// assert
AssertEquals_BOOL(Expected := TRUE, Actual := terminal_2.Channel1, Message := 'Channel1 follows SafeOut1');
AssertEquals_BOOL(Expected := FALSE, Actual := terminal_2.Channel2, Message := 'Channel2 follows SafeOut2');

// act: swap
group_2(Run := TRUE);
terminal_2(SafeOut1 := FALSE, SafeOut2 := TRUE, StartupTime := T#0S);

// assert
AssertEquals_BOOL(Expected := FALSE, Actual := terminal_2.Channel1, Message := 'Channel1 swapped');
AssertEquals_BOOL(Expected := TRUE, Actual := terminal_2.Channel2, Message := 'Channel2 swapped');
TEST_FINISHED_NAMED(__POUNAME());
END_METHOD

METHOD PRIVATE Test_ComErrorForcesChannelsFalse
TcUnit.TEST(__POUNAME());

// arrange: in Data with both outputs on
FOR i_3 := 1 TO 5 DO
    group_3(Run := TRUE);
    terminal_3(SafeOut1 := TRUE, SafeOut2 := TRUE, StartupTime := T#0S);
END_FOR
AssertEquals_BOOL(Expected := TRUE, Actual := terminal_3.Channel2, Message := 'Channel2 on before the error');

// act
group_3(Run := TRUE);
terminal_3(SafeOut1 := TRUE, SafeOut2 := TRUE, InjectComError := TRUE, StartupTime := T#0S);

// assert
AssertEquals_BOOL(Expected := TRUE, Actual := terminal_3.ComError, Message := 'com error');
AssertEquals_BOOL(Expected := FALSE, Actual := terminal_3.Channel1, Message := 'Channel1 fail-safe on com error');
AssertEquals_BOOL(Expected := FALSE, Actual := terminal_3.Channel2, Message := 'Channel2 fail-safe on com error');
TEST_FINISHED_NAMED(__POUNAME());
END_METHOD

METHOD PRIVATE Test_RegistersAsConnection
TcUnit.TEST(__POUNAME());

// act
group_4(Run := TRUE);
terminal_4(StartupTime := T#0S);

// assert
AssertEquals_UINT(Expected := 1, Actual := group_4.ConnectionCount, Message := 'one connection registered');
AssertEquals_UINT(Expected := 0, Actual := group_4.FunctionBlockCount, Message := 'no function blocks');
TEST_FINISHED_NAMED(__POUNAME());
END_METHOD

METHOD PRIVATE Test_GroupNotRunningForcesChannelsFalse
TcUnit.TEST(__POUNAME());
// arrange: connection in Data with the group running
FOR i_5 := 1 TO 10 DO
    group_5(Run := TRUE, ModuleFault := FALSE);
    terminal_5(StartupTime := T#0S, SafeOut1 := TRUE, SafeOut2 := TRUE);
END_FOR
AssertEquals_BOOL(Expected := TRUE, Actual := terminal_5.Channel1, Message := 'channel on while the group runs');
// act: group STOP (the connection stays in Data)
group_5(Run := FALSE, ModuleFault := FALSE);
terminal_5(StartupTime := T#0S, SafeOut1 := TRUE, SafeOut2 := TRUE);
// assert
AssertEquals_BOOL(Expected := TRUE, Actual := terminal_5.InDataState, Message := 'still in Data');
AssertEquals_BOOL(Expected := FALSE, Actual := terminal_5.Channel1, Message := 'outputs off with the group in STOP');
// act: group ERROR
group_5(Run := TRUE, ModuleFault := TRUE);
terminal_5(StartupTime := T#0S, SafeOut1 := TRUE, SafeOut2 := TRUE);
group_5(Run := TRUE, ModuleFault := TRUE);
terminal_5(StartupTime := T#0S, SafeOut1 := TRUE, SafeOut2 := TRUE);
AssertEquals_BYTE(Expected := TO_BYTE(E_SafeGroupState.Error), Actual := group_5.State, Message := 'group in ERROR');
AssertEquals_BOOL(Expected := FALSE, Actual := terminal_5.Channel2, Message := 'outputs off with the group in ERROR');
TEST_FINISHED_NAMED(__POUNAME());
END_METHOD

END_FUNCTION_BLOCK

// ---- Core/T_SafeOutputTerminal2.TcPOU
// Model of a two channel safe output terminal (EL2912): a TwinSAFE connection with two channels.
// Declare it in its group:  outputTerminal : T_SafeOutputTerminal2(group := safetyGroup);
// SafeOut1..2 are wired from FB outputs; Channel1..2 are the simulated field outputs,
// forced FALSE (fail-safe) unless the connection is in the Data state and the group is in RUN (OutputsEnabled).
FUNCTION_BLOCK T_SafeOutputTerminal2 EXTENDS T_SafeConnection
VAR_INPUT
    SafeOut1 : BOOL;
    SafeOut2 : BOOL;
END_VAR
VAR_OUTPUT
    Channel1 : BOOL;
    Channel2 : BOOL;
END_VAR

SUPER^();
Channel1 := SafeOut1 AND OutputsEnabled;
Channel2 := SafeOut2 AND OutputsEnabled;

END_FUNCTION_BLOCK

// ---- Tests/T_SafeConnShutdown_Tests.TcPOU
FUNCTION_BLOCK T_SafeConnShutdown_Tests EXTENDS TcUnit.FB_TestSuite
VAR
    // Test_DeactivateShutsDownConnection
    group_1 : T_SafeGroup;
    conn_1 : T_SafeConnection(group := group_1);
    fb_1 : T_SafeConnShutdown(group := group_1, connection := conn_1);
    i_1 : INT;
END_VAR

Test_DeactivateShutsDownConnection();

METHOD PRIVATE Test_DeactivateShutsDownConnection
TcUnit.TEST(__POUNAME());

// arrange: connection up
FOR i_1 := 1 TO 5 DO
    group_1(Run := TRUE);
    conn_1(StartupTime := T#0S);
    fb_1(Deactivate1 := FALSE);
END_FOR

AssertEquals_BOOL(Expected := FALSE, Actual := fb_1.Deactivated, Message := 'connection up');
// act
group_1(Run := TRUE);
fb_1(Deactivate1 := TRUE);
conn_1(StartupTime := T#0S);
fb_1(Deactivate1 := TRUE);
// assert
AssertEquals_BOOL(Expected := TRUE, Actual := conn_1.IsShutdown, Message := 'connection shut down');
AssertEquals_BOOL(Expected := TRUE, Actual := fb_1.Deactivated, Message := 'Deactivated output on');

// act: release
FOR i_1 := 1 TO 6 DO
    group_1(Run := TRUE);
    fb_1(Deactivate1 := FALSE);
    conn_1(StartupTime := T#0S);
END_FOR

AssertEquals_BOOL(Expected := TRUE, Actual := conn_1.InDataState, Message := 'connection re-established');
AssertEquals_BOOL(Expected := FALSE, Actual := fb_1.Deactivated, Message := 'Deactivated output off');
TEST_FINISHED_NAMED(__POUNAME());
END_METHOD

END_FUNCTION_BLOCK

// ---- FunctionBlocks/T_SafeConnShutdown.TcPOU
// Model of the TwinSAFE FB CONNECTION SHUTDOWN.
// Shuts down the assigned connection while the Deactivate inputs are TRUE and reports Deactivated
// once the connection is shut down (also when the partner shut it down). The connection is assigned
// at construction (the Connection ID of the Safety Editor):
//     connShutdown : T_SafeConnShutdown(group := safetyGroup, connection := toolConnection);
{attribute 'reflection'}
FUNCTION_BLOCK T_SafeConnShutdown EXTENDS T_SafeFunctionBlockBase
VAR_INPUT
    Deactivate1 : BOOL;
    Deactivate2 : BOOL;
    Parameters : ST_SafeConnShutdownParameters;
END_VAR
VAR_OUTPUT
    Deactivated : BOOL;
END_VAR
VAR
    {attribute 'is_connected' := 'Deactivate1'}
    _deactivate1Connected : BOOL;
    {attribute 'is_connected' := 'Deactivate2'}
    _deactivate2Connected : BOOL;
    _connection : REFERENCE TO T_SafeConnection;
    _pairs : ARRAY[1..1] OF T_SafeInputPair;
    _state : E_SafeFbState := E_SafeFbState.Stop;
    _prevState : E_SafeFbState;
END_VAR

SUPER^();

PROPERTY ConnShutdownState : E_SafeFbState
GET
ConnShutdownState := _state;
END_GET
END_PROPERTY

METHOD FB_init : BOOL
VAR_INPUT
    bInitRetains : BOOL;
    bInCopyCode : BOOL;
    group : REFERENCE TO T_SafeGroup; // the TwinSAFE group this block belongs to
    connection : REFERENCE TO T_SafeConnection; // the connection to shut down (Connection ID)
END_VAR
// the base FB_init (group registration) is called implicitly by TwinCAT
_connection REF= connection;
END_METHOD

METHOD PROTECTED Process
VAR
    acknowledge : BOOL;
    deactivate : BOOL;
    operating : BOOL;
    stateBefore : E_SafeFbState;
    passes : USINT;
END_VAR
acknowledge := (_state = E_SafeFbState.Error) AND _errAck;
_pairs[1](
    In1 := Deactivate1,
    In2 := Deactivate2,
    Active1 := _deactivate1Connected,
    Active2 := _deactivate2Connected,
    MakeContact1 := Parameters.Deactivate1MakeContact,
    MakeContact2 := Parameters.Deactivate2MakeContact,
    DiscrepancyTime := Parameters.DiscrepancyTime,
    Monitor := _fbRun,
    SafeInputsAfterDiscError := Parameters.SafeInputsAfterDiscError,
    Acknowledge := acknowledge
);

deactivate := _pairs[1].IsActive AND _pairs[1].AllTrue;

IF NOT _fbRun AND _state <> E_SafeFbState.Error AND _state <> E_SafeFbState.Reset THEN
    _state := E_SafeFbState.Stop;
END_IF

operating := (_state = E_SafeFbState.Safe) OR (_state = E_SafeFbState.Run);

IF _pairs[1].DiscrepancyError AND operating THEN
    UpdateDiscrepancyDiag();
    _state := E_SafeFbState.Error;
END_IF

passes := 0;

REPEAT
    stateBefore := _state;

    CASE _state OF
        E_SafeFbState.Stop:
            IF StateChanged() THEN
                Deactivated := FALSE;
                Error       := FALSE;
                Diag        := 0;
            END_IF

            _connection.LocalShutdown := FALSE;

            IF _fbRun THEN
                _state := E_SafeFbState.Safe;
            END_IF

        E_SafeFbState.Safe:
            IF StateChanged() THEN
                Deactivated := FALSE;
            END_IF

            _connection.LocalShutdown := deactivate;

            IF _connection.IsShutdown THEN
                _state := E_SafeFbState.Run;
            END_IF

        E_SafeFbState.Run:
            IF StateChanged() THEN
                Deactivated := TRUE;
            END_IF

            _connection.LocalShutdown := deactivate;

            IF NOT _connection.IsShutdown THEN
                _state := E_SafeFbState.Safe;
            END_IF

        E_SafeFbState.Error:
            IF StateChanged() THEN
                Deactivated := FALSE;
                Error       := TRUE;
            END_IF

            _connection.LocalShutdown := FALSE;
            UpdateDiscrepancyDiag();

            IF _errAck AND NOT _pairs[1].DiscrepancyError THEN
                _state := E_SafeFbState.Reset;
            END_IF

        E_SafeFbState.Reset:
            IF StateChanged() THEN
                Error := FALSE;
                Diag  := 0;
            END_IF

            IF _errAckFallingEdge THEN
                _state := SEL(_fbRun, E_SafeFbState.Stop, E_SafeFbState.Safe);
            END_IF
    END_CASE

    passes := passes + 1;
UNTIL (stateBefore = _state) OR (passes >= 3)
END_REPEAT

State := TO_BYTE(_state);
END_METHOD

METHOD PRIVATE StateChanged : BOOL
IF _prevState = _state THEN
    RETURN;
END_IF

_prevState   := _state;
StateChanged := TRUE;
END_METHOD

// Mirrors the discrepancy state of every pair into the diagnostic bits.
METHOD PRIVATE UpdateDiscrepancyDiag
VAR
    i : USINT;
END_VAR
FOR i := 1 TO 1 DO
    IF _pairs[i].DiscrepancyError THEN
        SetDiagBit(0);

        IF _pairs[i].AwaitingSafeInputs THEN
            SetDiagBit(8);
        ELSE
            ClearDiagBit(8);
        END_IF
    END_IF
END_FOR
END_METHOD

END_FUNCTION_BLOCK

// ---- Tests/T_SafeGroup_Tests.TcPOU
FUNCTION_BLOCK T_SafeGroup_Tests EXTENDS TcUnit.FB_TestSuite
VAR
    // Test_StopWhenRunFalse
    group_1 : T_SafeGroup;
    fb_1 : T_SafeAnd(group := group_1);
    // Test_RunsFunctionBlocksWithoutConnections
    group_2 : T_SafeGroup;
    fb_2 : T_SafeAnd(group := group_2);
    // Test_FbErrorStopsGroupAndErrAckRecovers
    group_3 : T_SafeGroup;
    eStop_3 : T_SafeEStop(group := group_3);
    andFb_3 : T_SafeAnd(group := group_3);
    // Test_ConnectionStartupAndComError
    group_4 : T_SafeGroup;
    terminal_4 : T_SafeInputTerminal(group := group_4);
    state_4 : INT := 10;
    waitTimer_4 : TON;
    // Test_RegistersMoreThanSixtyFourBlocks
    group_5 : T_SafeGroup;
    blocks_5 : ARRAY[1..70] OF T_SafeAnd(group := group_5);
    // Test_RefusesTheSixtyFifthConnection
    group_6 : T_SafeGroup;
    terminals_6 : ARRAY[1..65] OF T_SafeInputTerminal(group := group_6);
END_VAR

Test_StopWhenRunFalse();
Test_RunsFunctionBlocksWithoutConnections();
Test_FbErrorStopsGroupAndErrAckRecovers();
Test_ConnectionStartupAndComError();
Test_RegistersMoreThanSixtyFourBlocks();
Test_RefusesTheSixtyFifthConnection();

METHOD PRIVATE Test_ConnectionStartupAndComError
TcUnit.TEST(__POUNAME());
waitTimer_4();

CASE state_4 OF
    10:
        // arrange: terminal_4 starting up
        group_4(Run := TRUE, ErrAck := FALSE);
        terminal_4(InjectComError := FALSE, StartupTime := T#150MS);
        group_4(Run := TRUE, ErrAck := FALSE);
        terminal_4(InjectComError := FALSE, StartupTime := T#150MS);
        // assert
        AssertEquals_BYTE(
            Expected := TO_BYTE(E_SafeGroupState.Start),
            Actual := group_4.State,
            Message := 'group START while the connection starts up'
        );

        AssertEquals_BOOL(Expected := TRUE, Actual := group_4.ComStartup, Message := 'ComStartup');
        state_4 := 20;
        waitTimer_4(IN := TRUE, PT := T#400MS);
    20:
        group_4(Run := TRUE, ErrAck := FALSE);
        terminal_4(InjectComError := FALSE, StartupTime := T#150MS);

        IF NOT waitTimer_4.Q THEN
            RETURN;
        END_IF

        waitTimer_4(IN := FALSE);
        AssertEquals_BYTE(Expected := TO_BYTE(E_SafeGroupState.Run), Actual := group_4.State, Message := 'group RUN once the connection is in Data');
        // act: communication error
        group_4(Run := TRUE, ErrAck := FALSE);
        terminal_4(InjectComError := TRUE, StartupTime := T#150MS);
        group_4(Run := TRUE, ErrAck := FALSE);
        terminal_4(InjectComError := FALSE, StartupTime := T#150MS);
        AssertEquals_BOOL(Expected := TRUE, Actual := group_4.ComErr, Message := 'ComErr');
        AssertEquals_BYTE(Expected := TO_BYTE(E_SafeGroupState.Error), Actual := group_4.State, Message := 'group ERROR');
        group_4(Run := TRUE, ErrAck := TRUE);
        terminal_4(InjectComError := FALSE, StartupTime := T#150MS);
        group_4(Run := TRUE, ErrAck := TRUE);
        terminal_4(InjectComError := FALSE, StartupTime := T#150MS);
        AssertEquals_BYTE(Expected := TO_BYTE(E_SafeGroupState.Reset), Actual := group_4.State, Message := 'group RESET');
        group_4(Run := TRUE, ErrAck := FALSE);
        terminal_4(InjectComError := FALSE, StartupTime := T#150MS);
        AssertEquals_BYTE(Expected := TO_BYTE(E_SafeGroupState.Start), Actual := group_4.State, Message := 'group START again after ack');
        state_4 := 30;
        waitTimer_4(IN := TRUE, PT := T#400MS);
    30:
        group_4(Run := TRUE, ErrAck := FALSE);
        terminal_4(InjectComError := FALSE, StartupTime := T#150MS);

        IF NOT waitTimer_4.Q THEN
            RETURN;
        END_IF

        waitTimer_4(IN := FALSE);
        AssertEquals_BYTE(Expected := TO_BYTE(E_SafeGroupState.Run), Actual := group_4.State, Message := 'group RUN after reconnection');
        TEST_FINISHED_NAMED(__POUNAME());
        state_4 := 10;
END_CASE
END_METHOD

METHOD PRIVATE Test_FbErrorStopsGroupAndErrAckRecovers
TcUnit.TEST(__POUNAME());
// arrange: an AND that runs and an ESTOP that will raise an EDM error
group_3(Run := TRUE, ErrAck := FALSE);
eStop_3(Restart := FALSE, EDM1 := FALSE, EStopIn1 := TRUE);
andFb_3(AndIn1 := TRUE, AndIn2 := TRUE);
group_3(Run := TRUE, ErrAck := FALSE);
eStop_3(Restart := FALSE, EDM1 := FALSE, EStopIn1 := TRUE);
andFb_3(AndIn1 := TRUE, AndIn2 := TRUE);
AssertEquals_BOOL(Expected := TRUE, Actual := andFb_3.AndOut, Message := 'AND running before the error');
// act: restart with missing feedback -> FB error
group_3(Run := TRUE, ErrAck := FALSE);
eStop_3(Restart := TRUE, EDM1 := FALSE, EStopIn1 := TRUE);
andFb_3(AndIn1 := TRUE, AndIn2 := TRUE);
group_3(Run := TRUE, ErrAck := FALSE);
eStop_3(Restart := FALSE, EDM1 := FALSE, EStopIn1 := TRUE);
andFb_3(AndIn1 := TRUE, AndIn2 := TRUE);
// assert
AssertEquals_BOOL(Expected := TRUE, Actual := group_3.FbErr, Message := 'FbErr');
AssertEquals_BYTE(Expected := TO_BYTE(E_SafeGroupState.Error), Actual := group_3.State, Message := 'group ERROR');
AssertEquals_BYTE(Expected := TO_BYTE(E_SafeGroupDiag.FbError), Actual := group_3.Diag, Message := 'group diag FBERROR');
AssertEquals_BOOL(Expected := FALSE, Actual := andFb_3.AndOut, Message := 'other FB outputs forced safe');
AssertEquals_BYTE(Expected := TO_BYTE(E_SafeFbState.Stop), Actual := andFb_3.State, Message := 'other FB STOP');
// act: ErrAck 0 -> 1 -> 0
group_3(Run := TRUE, ErrAck := TRUE);
eStop_3(Restart := FALSE, EDM1 := FALSE, EStopIn1 := TRUE);
andFb_3(AndIn1 := TRUE, AndIn2 := TRUE);
group_3(Run := TRUE, ErrAck := TRUE);
eStop_3(Restart := FALSE, EDM1 := FALSE, EStopIn1 := TRUE);
andFb_3(AndIn1 := TRUE, AndIn2 := TRUE);
AssertEquals_BYTE(Expected := TO_BYTE(E_SafeGroupState.Reset), Actual := group_3.State, Message := 'group RESET while ErrAck 1');
group_3(Run := TRUE, ErrAck := FALSE);
eStop_3(Restart := FALSE, EDM1 := FALSE, EStopIn1 := TRUE);
andFb_3(AndIn1 := TRUE, AndIn2 := TRUE);
group_3(Run := TRUE, ErrAck := FALSE);
eStop_3(Restart := FALSE, EDM1 := FALSE, EStopIn1 := TRUE);
andFb_3(AndIn1 := TRUE, AndIn2 := TRUE);
AssertEquals_BYTE(Expected := TO_BYTE(E_SafeGroupState.Run), Actual := group_3.State, Message := 'group RUN after ErrAck');
AssertEquals_BOOL(Expected := TRUE, Actual := andFb_3.AndOut, Message := 'AND running again');
AssertEquals_BYTE(Expected := TO_BYTE(E_SafeFbState.Safe), Actual := eStop_3.State, Message := 'ESTOP back in SAFE awaiting restart');
TEST_FINISHED_NAMED(__POUNAME());
END_METHOD

METHOD PRIVATE Test_RunsFunctionBlocksWithoutConnections
TcUnit.TEST(__POUNAME());
// act
group_2(Run := TRUE);
fb_2(AndIn1 := TRUE, AndIn2 := TRUE);
group_2(Run := TRUE);
fb_2(AndIn1 := TRUE, AndIn2 := TRUE);
// assert
AssertEquals_BYTE(Expected := TO_BYTE(E_SafeGroupState.Run), Actual := group_2.State, Message := 'group RUN');
AssertEquals_BOOL(Expected := TRUE, Actual := fb_2.AndOut, Message := 'FB executed');
AssertEquals_BOOL(Expected := TRUE, Actual := group_2.FbRun, Message := 'all FBs running');
TEST_FINISHED_NAMED(__POUNAME());
END_METHOD

METHOD PRIVATE Test_StopWhenRunFalse
TcUnit.TEST(__POUNAME());
// act
group_1(Run := FALSE);
fb_1(AndIn1 := TRUE, AndIn2 := TRUE);
// assert
AssertEquals_BYTE(Expected := TO_BYTE(E_SafeGroupState.Stop), Actual := group_1.State, Message := 'group STOP');
AssertEquals_BYTE(Expected := TO_BYTE(E_SafeFbState.Stop), Actual := fb_1.State, Message := 'FB STOP');
AssertEquals_BOOL(Expected := FALSE, Actual := group_1.InRun, Message := 'InRun off');
TEST_FINISHED_NAMED(__POUNAME());
END_METHOD

METHOD PRIVATE Test_RegistersMoreThanSixtyFourBlocks
TcUnit.TEST(__POUNAME());
// arrange: 70 blocks joined group_5 at initialisation
// assert
AssertEquals_UINT(Expected := 70, Actual := group_5.FunctionBlockCount, Message := 'every block registered');
AssertEquals_BOOL(Expected := FALSE, Actual := group_5.RegistrationRefused, Message := 'none refused');
TEST_FINISHED_NAMED(__POUNAME());
END_METHOD

METHOD PRIVATE Test_RefusesTheSixtyFifthConnection
TcUnit.TEST(__POUNAME());
// arrange: 65 terminals tried to join group_6 at initialisation
// assert
AssertEquals_UINT(Expected := 64, Actual := group_6.ConnectionCount, Message := 'the cap holds');
AssertEquals_BOOL(Expected := TRUE, Actual := group_6.RegistrationRefused, Message := 'the refusal is visible');
TEST_FINISHED_NAMED(__POUNAME());
END_METHOD

END_FUNCTION_BLOCK

// ---- Core/T_SafeInputTerminal.TcPOU
// Model of a four channel safe input terminal (EL1904): a TwinSAFE connection with four channels.
// Declare it in its group:  inputTerminal : T_SafeInputTerminal(group := safetyGroup);
// Channel1..4 are the simulated field signals; SafeIn1..4 are what the TwinSAFE logic sees:
// forced FALSE (fail-safe) unless the connection is in the Data state.
FUNCTION_BLOCK T_SafeInputTerminal EXTENDS T_SafeConnection
VAR_INPUT
    Channel1 : BOOL;
    Channel2 : BOOL;
    Channel3 : BOOL;
    Channel4 : BOOL;
END_VAR
VAR_OUTPUT
    SafeIn1 : BOOL;
    SafeIn2 : BOOL;
    SafeIn3 : BOOL;
    SafeIn4 : BOOL;
END_VAR

SUPER^();
SafeIn1 := Channel1 AND InDataState;
SafeIn2 := Channel2 AND InDataState;
SafeIn3 := Channel3 AND InDataState;
SafeIn4 := Channel4 AND InDataState;

END_FUNCTION_BLOCK

// ---- Tests/User_FB_Tests/T_SafePulse_UserFB_Tests.TcPOU
// Tests of the example user FB T_SafePulse_UserFB: TonOut is a pulse of DelayTime while TonIn1 is held.
FUNCTION_BLOCK T_SafePulse_UserFB_Tests EXTENDS TcUnit.FB_TestSuite
VAR
    // Test_PulseForDelayTimeWhileInputHeld
    group_1 : T_SafeGroup;
    fb_1 : T_SafePulse_UserFB(group := group_1) := (Parameters := (DelayTime := T#100MS));
    state_1 : INT := 10;
    waitTimer_1 : TON;
    // Test_PulseEndsWhenInputDrops
    group_2 : T_SafeGroup;
    fb_2 : T_SafePulse_UserFB(group := group_2) := (Parameters := (DelayTime := T#100MS));
    // Test_StoppedGivesNoOutput
    group_3 : T_SafeGroup;
    fb_3 : T_SafePulse_UserFB(group := group_3) := (Parameters := (DelayTime := T#100MS));
    // Test_InnerBlocksJoinTheGroup
    group_4 : T_SafeGroup;
    fb_4 : T_SafePulse_UserFB(group := group_4);
END_VAR

Test_PulseForDelayTimeWhileInputHeld();
Test_PulseEndsWhenInputDrops();
Test_StoppedGivesNoOutput();
Test_InnerBlocksJoinTheGroup();

METHOD PRIVATE Test_InnerBlocksJoinTheGroup
TcUnit.TEST(__POUNAME());
// assert: the composite registered itself and passed the group on to its TON and AND
AssertEquals_UINT(Expected := 3, Actual := group_4.FunctionBlockCount, Message := 'composite and its two inner blocks registered');
TEST_FINISHED_NAMED(__POUNAME());
END_METHOD

METHOD PRIVATE Test_PulseEndsWhenInputDrops
TcUnit.TEST(__POUNAME());
// act / assert
group_2(Run := TRUE);
fb_2(TonIn1 := TRUE);
AssertEquals_BOOL(Expected := TRUE, Actual := fb_2.TonOut, Message := 'pulse on');
AssertEquals_BOOL(Expected := TRUE, Actual := fb_2.IsRunning, Message := 'reports Run to the group while it runs');
fb_2(TonIn1 := FALSE);
AssertEquals_BOOL(Expected := FALSE, Actual := fb_2.TonOut, Message := 'pulse cut off when the input drops');
TEST_FINISHED_NAMED(__POUNAME());
END_METHOD

METHOD PRIVATE Test_PulseForDelayTimeWhileInputHeld
TcUnit.TEST(__POUNAME());
waitTimer_1();

CASE state_1 OF
    10:
        // act: input on, the pulse starts
        group_1(Run := TRUE);
        fb_1(TonIn1 := TRUE);
        // assert
        AssertEquals_BOOL(Expected := TRUE, Actual := fb_1.TonOut, Message := 'pulse starts with the input');
        state_1 := 20;
        waitTimer_1(IN := TRUE, PT := T#50MS);
    20:
        group_1(Run := TRUE);
        fb_1(TonIn1 := TRUE);

        IF NOT waitTimer_1.Q THEN
            RETURN;
        END_IF

        waitTimer_1(IN := FALSE);
        // assert: still inside the delay time
        AssertEquals_BOOL(Expected := TRUE, Actual := fb_1.TonOut, Message := 'pulse still on inside the delay time');
        state_1 := 30;
        waitTimer_1(IN := TRUE, PT := T#200MS);
    30:
        group_1(Run := TRUE);
        fb_1(TonIn1 := TRUE);

        IF NOT waitTimer_1.Q THEN
            RETURN;
        END_IF

        waitTimer_1(IN := FALSE);
        // assert: the delay has elapsed, the pulse is over although the input is still held
        AssertEquals_BOOL(Expected := FALSE, Actual := fb_1.TonOut, Message := 'pulse ends after the delay time');
        // act: release and re-apply the input
        fb_1(TonIn1 := FALSE);
        AssertEquals_BOOL(Expected := FALSE, Actual := fb_1.TonOut, Message := 'no output with the input off');
        fb_1(TonIn1 := TRUE);
        AssertEquals_BOOL(Expected := TRUE, Actual := fb_1.TonOut, Message := 'a new pulse starts on the next rising edge');
        TEST_FINISHED_NAMED(__POUNAME());
        state_1 := 10;
END_CASE
END_METHOD

METHOD PRIVATE Test_StoppedGivesNoOutput
TcUnit.TEST(__POUNAME());
// act
group_3(Run := FALSE);
fb_3(TonIn1 := TRUE);
// assert
AssertEquals_BOOL(Expected := FALSE, Actual := fb_3.TonOut, Message := 'no output while the group is stopped');
AssertEquals_BOOL(Expected := FALSE, Actual := fb_3.IsRunning, Message := 'not running while the group is stopped');
TEST_FINISHED_NAMED(__POUNAME());
END_METHOD

END_FUNCTION_BLOCK

// ---- Examples/Example_UserFbs/T_SafePulse_UserFB.TcPOU
FUNCTION_BLOCK T_SafePulse_UserFB EXTENDS T_SafeFunctionBlockBase
VAR_INPUT
	TonIn1 : BOOL;
	Parameters : ST_SafeTimerParameters;
END_VAR
VAR_OUTPUT
	TonOut : BOOL;
END_VAR
VAR
	safeTon : T_SafeTon(_group);
	safeAnd : T_SafeAnd(_group);
END_VAR

SUPER^();

METHOD FB_init : BOOL
VAR_INPUT
	bInitRetains	: BOOL;
	bInCopyCode	: BOOL;
	group	: REFERENCE TO T_SafeGroup;
END_VAR
safeAnd.SetGroupReference(bInCopyCode := bInCopyCode, group := group);
safeTon.SetGroupReference(bInCopyCode := bInCopyCode, group := group);
END_METHOD

METHOD PROTECTED Process
safeTon(TonIn1 := TonIn1, Parameters := Parameters); // T_SafeTon
safeAnd(AndIn1 := NOT safeTon.TonOut, AndIn2 := TonIn1); // T_SafeAnd
TonOut := safeAnd.AndOut;
END_METHOD

END_FUNCTION_BLOCK

// ---- Tests/User_FB_Tests/T_SafeRTrig_UserFB_Tests.TcPOU
// Tests of the example user FB T_SafeRTrig_UserFB: Trigger is on for one cycle on the rising edge of Signal.
FUNCTION_BLOCK T_SafeRTrig_UserFB_Tests EXTENDS TcUnit.FB_TestSuite
VAR
    // Test_TriggerForOneCycleOnRisingEdge
    group_1 : T_SafeGroup;
    fb_1 : T_SafeRTrig_UserFB(group := group_1);
    // Test_StoppedGivesNoOutput
    group_2 : T_SafeGroup;
    fb_2 : T_SafeRTrig_UserFB(group := group_2);
    // Test_InnerBlocksJoinTheGroup
    group_3 : T_SafeGroup;
    fb_3 : T_SafeRTrig_UserFB(group := group_3);
END_VAR

Test_TriggerForOneCycleOnRisingEdge();
Test_StoppedGivesNoOutput();
Test_InnerBlocksJoinTheGroup();

METHOD PRIVATE Test_InnerBlocksJoinTheGroup
TcUnit.TEST(__POUNAME());
// assert: the composite registered itself and passed the group on to its RS and AND
AssertEquals_UINT(Expected := 3, Actual := group_3.FunctionBlockCount, Message := 'composite and its two inner blocks registered');
TEST_FINISHED_NAMED(__POUNAME());
END_METHOD

METHOD PRIVATE Test_StoppedGivesNoOutput
TcUnit.TEST(__POUNAME());
// act
group_2(Run := FALSE);
fb_2(Signal := TRUE);
// assert
AssertEquals_BOOL(Expected := FALSE, Actual := fb_2.Trigger, Message := 'no output while the group is stopped');
AssertEquals_BOOL(Expected := FALSE, Actual := fb_2.IsRunning, Message := 'not running while the group is stopped');
TEST_FINISHED_NAMED(__POUNAME());
END_METHOD

METHOD PRIVATE Test_TriggerForOneCycleOnRisingEdge
TcUnit.TEST(__POUNAME());
// act / assert
group_1(Run := TRUE);
fb_1(Signal := FALSE);
AssertEquals_BOOL(Expected := FALSE, Actual := fb_1.Trigger, Message := 'no trigger while the signal is off');
AssertEquals_BOOL(Expected := TRUE, Actual := fb_1.IsRunning, Message := 'reports Run to the group while it runs');
fb_1(Signal := TRUE);
AssertEquals_BOOL(Expected := TRUE, Actual := fb_1.Trigger, Message := 'trigger on the rising edge');
fb_1(Signal := TRUE);
AssertEquals_BOOL(Expected := FALSE, Actual := fb_1.Trigger, Message := 'trigger lasts one cycle');
fb_1(Signal := FALSE);
AssertEquals_BOOL(Expected := FALSE, Actual := fb_1.Trigger, Message := 'no trigger on the falling edge');
fb_1(Signal := TRUE);
AssertEquals_BOOL(Expected := TRUE, Actual := fb_1.Trigger, Message := 'triggers again on the next rising edge');
TEST_FINISHED_NAMED(__POUNAME());
END_METHOD

END_FUNCTION_BLOCK

// ---- Examples/Example_UserFbs/T_SafeRTrig_UserFB.TcPOU
FUNCTION_BLOCK T_SafeRTrig_UserFB EXTENDS T_SafeFunctionBlockBase
VAR_INPUT
	Signal : BOOL;
END_VAR
VAR_OUTPUT
	Trigger : BOOL;
END_VAR
VAR
	safeRs : T_SafeRs(_group);
	safeAnd : T_SafeAnd(_group);
END_VAR

SUPER^();

METHOD FB_init : BOOL
VAR_INPUT
	bInitRetains	: BOOL;
	bInCopyCode	: BOOL;
	group	: REFERENCE TO T_SafeGroup;
END_VAR
safeRs.SetGroupReference(bInCopyCode := bInCopyCode, group := group);
safeAnd.SetGroupReference(bInCopyCode := bInCopyCode, group := group);
END_METHOD

METHOD PROTECTED Process
safeAnd(AndIn1 := Signal, AndIn2 := NOT safeRs.RsOut); // T_SafeAnd
safeRs(Set := Signal, Reset := NOT Signal); // T_SafeRs
Trigger := safeAnd.AndOut;
END_METHOD

END_FUNCTION_BLOCK

// ---- Tests/T_SafeAnd_Tests_CFC.TcPOU
    // CFC twin of T_SafeAnd_Tests: the same tests drawn as CFC diagrams, the way a TwinSAFE project is authored.
    FUNCTION_BLOCK T_SafeAnd_Tests_CFC EXTENDS T_SafeCfcTestSuite
    VAR
    // Test_AllConnectedInputsTrueGivesRun
    group_1 : T_SafeGroup;
    fb_1 : T_SafeAnd(group := group_1);
    // Test_OneInputFalseGivesSafe
    group_2 : T_SafeGroup;
    fb_2 : T_SafeAnd(group := group_2);
    // Test_UnconnectedInputsIgnoredAndMakeContactNegated
    group_3 : T_SafeGroup;
    fb_3 : T_SafeAnd(group := group_3) := (Parameters := (In2MakeContact := TRUE));
    // Test_StoppedGivesNoOutput
    group_4 : T_SafeGroup;
    fb_4 : T_SafeAnd(group := group_4);
END_VAR

Test_AllConnectedInputsTrueGivesRun();
Test_OneInputFalseGivesSafe();
Test_UnconnectedInputsIgnoredAndMakeContactNegated();
Test_StoppedGivesNoOutput();

METHOD PRIVATE Test_AllConnectedInputsTrueGivesRun
// note: this text did not pass the execution check against the stored diagram
StartTest(TestName := 'Test_AllConnectedInputsTrueGivesRun');
group_1(Run := TRUE, ErrAck := FALSE); // T_SafeGroup
fb_1(AndIn1 := TRUE, AndIn2 := TRUE); // T_SafeAnd
AssertEquals_BOOL(Expected := TRUE, Actual := fb_1.AndOut, Message := 'output on when all connected inputs are 1');
AssertEquals_BYTE(Expected := TO_BYTE(E_SafeFbState.Run), Actual := fb_1.State, Message := 'state RUN');
FinishTest(TestName := 'Test_AllConnectedInputsTrueGivesRun');
END_METHOD

METHOD PRIVATE Test_OneInputFalseGivesSafe
// note: this text did not pass the execution check against the stored diagram
StartTest(TestName := 'Test_OneInputFalseGivesSafe');
group_2(Run := TRUE, ErrAck := FALSE); // T_SafeGroup
fb_2(AndIn1 := TRUE, AndIn2 := FALSE); // T_SafeAnd
AssertEquals_BOOL(Expected := FALSE, Actual := fb_2.AndOut, Message := 'output off when a connected input is 0');
AssertEquals_BYTE(Expected := TO_BYTE(E_SafeFbState.Safe), Actual := fb_2.State, Message := 'state SAFE');
FinishTest(TestName := 'Test_OneInputFalseGivesSafe');
END_METHOD

METHOD PRIVATE Test_UnconnectedInputsIgnoredAndMakeContactNegated
// note: this text did not pass the execution check against the stored diagram
StartTest(TestName := 'Test_UnconnectedInputsIgnoredAndMakeContactNegated');
group_3(Run := TRUE, ErrAck := FALSE); // T_SafeGroup
fb_3(AndIn1 := TRUE, AndIn2 := FALSE); // T_SafeAnd
AssertEquals_BOOL(Expected := TRUE, Actual := fb_3.AndOut, Message := 'unconnected inputs ignored, make contact negated');
FinishTest(TestName := 'Test_UnconnectedInputsIgnoredAndMakeContactNegated');
END_METHOD

METHOD PRIVATE Test_StoppedGivesNoOutput
// note: this text did not pass the execution check against the stored diagram
StartTest(TestName := 'Test_StoppedGivesNoOutput');
group_4(Run := FALSE, ErrAck := FALSE); // T_SafeGroup
fb_4(AndIn1 := TRUE, AndIn2 := TRUE); // T_SafeAnd
AssertEquals_BOOL(Expected := FALSE, Actual := fb_4.AndOut, Message := 'no output while the group is stopped');
AssertEquals_BYTE(Expected := TO_BYTE(E_SafeFbState.Stop), Actual := fb_4.State, Message := 'state STOP');
FinishTest(TestName := 'Test_StoppedGivesNoOutput');
END_METHOD

END_FUNCTION_BLOCK

// ---- Tests/T_SafeCfcTestSuite.TcPOU
// Base of the CFC test suites. TcUnit's TEST and TEST_FINISHED_NAMED are functions without a return
// type, which a CFC box cannot call (the editor insists on a return pin), so the diagrams call these
// two methods instead. Everything else comes from TcUnit.FB_TestSuite.
FUNCTION_BLOCK ABSTRACT T_SafeCfcTestSuite EXTENDS TcUnit.FB_TestSuite

// Marks the start of a test (TcUnit.TEST). Call it first in every test method, every cycle.
METHOD PROTECTED StartTest
VAR_INPUT
    TestName : T_MaxString;
END_VAR
TcUnit.TEST(TestName);
END_METHOD

// Marks a test as finished (TcUnit.TEST_FINISHED_NAMED).
METHOD PROTECTED FinishTest
VAR_INPUT
    TestName : T_MaxString;
END_VAR
TcUnit.TEST_FINISHED_NAMED(TestName);
END_METHOD

END_FUNCTION_BLOCK

// ---- Tests/T_SafeInputPair_Tests_CFC.TcPOU
    // CFC twin of T_SafeInputPair_Tests: the same tests drawn as CFC diagrams, the way a TwinSAFE project is authored.
    FUNCTION_BLOCK T_SafeInputPair_Tests_CFC EXTENDS T_SafeCfcTestSuite
    VAR
    // Test_InactivePairNeverRequestsSafeState
    pair_1 : T_SafeInputPair;
    // Test_BreakContactRequestsSafeStateOnZero
    pair_2 : T_SafeInputPair;
    // Test_MakeContactRequestsSafeStateOnOne
    pair_3 : T_SafeInputPair;
    // Test_TwoChannelRequestsSafeStateIfEitherChannelLow
    pair_4 : T_SafeInputPair;
    // Test_DiscrepancyErrorAfterTimeoutAndResetAfterSafeInputs
    pair_5 : T_SafeInputPair;
    t1_5 : TON;
    t2_5 : TON;
    trig1_5 : R_TRIG;
    trig2_5 : R_TRIG;
END_VAR

Test_InactivePairNeverRequestsSafeState();
Test_BreakContactRequestsSafeStateOnZero();
Test_MakeContactRequestsSafeStateOnOne();
Test_TwoChannelRequestsSafeStateIfEitherChannelLow();
Test_DiscrepancyErrorAfterTimeoutAndResetAfterSafeInputs();

METHOD PRIVATE Test_InactivePairNeverRequestsSafeState
// note: this text did not pass the execution check against the stored diagram
StartTest(TestName := 'Test_InactivePairNeverRequestsSafeState');
pair_1(In1 := FALSE, In2 := FALSE, Active1 := FALSE, Active2 := FALSE, Monitor := TRUE); // T_SafeInputPair
AssertEquals_BOOL(Expected := FALSE, Actual := pair_1.SafeStateRequested, Message := 'inactive pair must not request the safe state');
AssertEquals_BOOL(Expected := FALSE, Actual := pair_1.IsActive, Message := 'pair should be inactive');
FinishTest(TestName := 'Test_InactivePairNeverRequestsSafeState');
END_METHOD

METHOD PRIVATE Test_BreakContactRequestsSafeStateOnZero
// note: this text did not pass the execution check against the stored diagram
StartTest(TestName := 'Test_BreakContactRequestsSafeStateOnZero');
pair_2(In1 := FALSE, Active1 := TRUE, Monitor := TRUE); // T_SafeInputPair
AssertEquals_BOOL(Expected := TRUE, Actual := pair_2.SafeStateRequested, Message := 'break contact at 0 must request the safe state');
pair_2(In1 := TRUE, Active1 := TRUE, Monitor := TRUE); // T_SafeInputPair
AssertEquals_BOOL(Expected := FALSE, Actual := pair_2.SafeStateRequested, Message := 'break contact at 1 must not request the safe state');
FinishTest(TestName := 'Test_BreakContactRequestsSafeStateOnZero');
END_METHOD

METHOD PRIVATE Test_MakeContactRequestsSafeStateOnOne
// note: this text did not pass the execution check against the stored diagram
StartTest(TestName := 'Test_MakeContactRequestsSafeStateOnOne');
pair_3(In1 := TRUE, Active1 := TRUE, MakeContact1 := TRUE, Monitor := TRUE); // T_SafeInputPair
AssertEquals_BOOL(Expected := TRUE, Actual := pair_3.SafeStateRequested, Message := 'make contact at 1 must request the safe state');
FinishTest(TestName := 'Test_MakeContactRequestsSafeStateOnOne');
END_METHOD

METHOD PRIVATE Test_TwoChannelRequestsSafeStateIfEitherChannelLow
// note: this text did not pass the execution check against the stored diagram
StartTest(TestName := 'Test_TwoChannelRequestsSafeStateIfEitherChannelLow');
pair_4(
    In1 := TRUE,
    In2 := FALSE,
    Active1 := TRUE,
    Active2 := TRUE,
    Monitor := TRUE,
    SafeInputsAfterDiscError := TRUE); // T_SafeInputPair
AssertEquals_BOOL(Expected := TRUE, Actual := pair_4.SafeStateRequested, Message := 'one low channel must request the safe state');
AssertEquals_BOOL(Expected := FALSE, Actual := pair_4.DiscrepancyError, Message := 'no discrepancy monitoring without a discrepancy time');
pair_4(
    In1 := TRUE,
    In2 := TRUE,
    Active1 := TRUE,
    Active2 := TRUE,
    Monitor := TRUE,
    SafeInputsAfterDiscError := TRUE); // T_SafeInputPair
AssertEquals_BOOL(Expected := FALSE, Actual := pair_4.SafeStateRequested, Message := 'both channels high must not request the safe state');
FinishTest(TestName := 'Test_TwoChannelRequestsSafeStateIfEitherChannelLow');
END_METHOD

METHOD PRIVATE Test_DiscrepancyErrorAfterTimeoutAndResetAfterSafeInputs
// note: this text did not pass the execution check against the stored diagram
StartTest(TestName := 'Test_DiscrepancyErrorAfterTimeoutAndResetAfterSafeInputs');
t1_5(IN := TRUE, PT := T#50MS); // TON
t2_5(IN := t1_5.Q, PT := T#200MS); // TON
trig1_5(CLK := t1_5.Q); // R_TRIG
trig2_5(CLK := t2_5.Q); // R_TRIG
pair_5(
    In1 := TRUE,
    In2 := FALSE,
    Active1 := TRUE,
    Active2 := TRUE,
    DiscrepancyTime := T#100MS,
    Monitor := TRUE,
    SafeInputsAfterDiscError := TRUE,
    Acknowledge := FALSE); // T_SafeInputPair
IF trig1_5.Q THEN AssertEquals_BOOL(Expected := FALSE, Actual := pair_5.DiscrepancyError, Message := 'no error before the discrepancy time'); END_IF
IF trig2_5.Q THEN AssertEquals_BOOL(Expected := TRUE, Actual := pair_5.DiscrepancyError, Message := 'error after the discrepancy time'); END_IF
IF trig2_5.Q THEN AssertEquals_BOOL(Expected := TRUE, Actual := pair_5.AwaitingSafeInputs, Message := 'error waits for both channels safe'); END_IF
IF trig2_5.Q THEN
    pair_5(
        In1 := TRUE,
        In2 := FALSE,
        Active1 := TRUE,
        Active2 := TRUE,
        DiscrepancyTime := T#100MS,
        Monitor := TRUE,
        SafeInputsAfterDiscError := TRUE,
        Acknowledge := TRUE); // T_SafeInputPair
END_IF
IF trig2_5.Q THEN AssertEquals_BOOL(Expected := TRUE, Actual := pair_5.DiscrepancyError, Message := 'acknowledge refused while a channel is still high'); END_IF
IF trig2_5.Q THEN
    pair_5(
        In1 := FALSE,
        In2 := FALSE,
        Active1 := TRUE,
        Active2 := TRUE,
        DiscrepancyTime := T#100MS,
        Monitor := TRUE,
        SafeInputsAfterDiscError := TRUE,
        Acknowledge := TRUE); // T_SafeInputPair
END_IF
IF trig2_5.Q THEN AssertEquals_BOOL(Expected := FALSE, Actual := pair_5.DiscrepancyError, Message := 'error cleared once both channels were safe'); END_IF
IF trig2_5.Q THEN FinishTest(TestName := 'Test_DiscrepancyErrorAfterTimeoutAndResetAfterSafeInputs'); END_IF
END_METHOD

END_FUNCTION_BLOCK

// ---- Tests/T_SafeOr_Tests_CFC.TcPOU
    // CFC twin of T_SafeOr_Tests: the same tests drawn as CFC diagrams, the way a TwinSAFE project is authored.
    FUNCTION_BLOCK T_SafeOr_Tests_CFC EXTENDS T_SafeCfcTestSuite
    VAR
    // Test_AnyConnectedInputTrueGivesRun
    group_1 : T_SafeGroup;
    fb_1 : T_SafeOr(group := group_1);
    // Test_AllFalseGivesSafe
    group_2 : T_SafeGroup;
    fb_2 : T_SafeOr(group := group_2);
END_VAR

Test_AnyConnectedInputTrueGivesRun();
Test_AllFalseGivesSafe();

METHOD PRIVATE Test_AnyConnectedInputTrueGivesRun
// note: this text did not pass the execution check against the stored diagram
StartTest(TestName := 'Test_AnyConnectedInputTrueGivesRun');
group_1(Run := TRUE, ErrAck := FALSE); // T_SafeGroup
fb_1(OrIn1 := FALSE, OrIn2 := TRUE); // T_SafeOr
AssertEquals_BOOL(Expected := TRUE, Actual := fb_1.OrOut, Message := 'output on when any connected input is 1');
FinishTest(TestName := 'Test_AnyConnectedInputTrueGivesRun');
END_METHOD

METHOD PRIVATE Test_AllFalseGivesSafe
// note: this text did not pass the execution check against the stored diagram
StartTest(TestName := 'Test_AllFalseGivesSafe');
group_2(Run := TRUE, ErrAck := FALSE); // T_SafeGroup
fb_2(OrIn1 := FALSE, OrIn2 := FALSE); // T_SafeOr
AssertEquals_BOOL(Expected := FALSE, Actual := fb_2.OrOut, Message := 'output off when all connected inputs are 0');
AssertEquals_BYTE(Expected := TO_BYTE(E_SafeFbState.Safe), Actual := fb_2.State, Message := 'state SAFE');
FinishTest(TestName := 'Test_AllFalseGivesSafe');
END_METHOD

END_FUNCTION_BLOCK

// ---- Tests/T_SafeXor_Tests_CFC.TcPOU
    // CFC twin of T_SafeXor_Tests: the same tests drawn as CFC diagrams, the way a TwinSAFE project is authored.
    FUNCTION_BLOCK T_SafeXor_Tests_CFC EXTENDS T_SafeCfcTestSuite
    VAR
    // Test_ConnectedPairsAreExclusiveOr
    group_1 : T_SafeGroup;
    fb_1 : T_SafeXor(group := group_1);
END_VAR

Test_ConnectedPairsAreExclusiveOr();

METHOD PRIVATE Test_ConnectedPairsAreExclusiveOr
// note: this text did not pass the execution check against the stored diagram
StartTest(TestName := 'Test_ConnectedPairsAreExclusiveOr');
group_1(Run := TRUE, ErrAck := FALSE); // T_SafeGroup
fb_1(Xor1In1 := TRUE, Xor2In1 := FALSE); // T_SafeXor
AssertEquals_BOOL(Expected := TRUE, Actual := fb_1.XorOut1, Message := 'connected pair 1 XOR');
AssertEquals_BOOL(Expected := FALSE, Actual := fb_1.XorOut2, Message := 'unconnected pair stays 0');
fb_1(Xor1In1 := TRUE, Xor2In1 := TRUE); // T_SafeXor
AssertEquals_BOOL(Expected := FALSE, Actual := fb_1.XorOut1, Message := 'both inputs 1 gives 0');
FinishTest(TestName := 'Test_ConnectedPairsAreExclusiveOr');
END_METHOD

END_FUNCTION_BLOCK

// ---- Tests/T_SafeDecouple_Tests_CFC.TcPOU
    // CFC twin of T_SafeDecouple_Tests: the same tests drawn as CFC diagrams, the way a TwinSAFE project is authored.
    FUNCTION_BLOCK T_SafeDecouple_Tests_CFC EXTENDS T_SafeCfcTestSuite
    VAR
    // Test_InputsLoopedToOutputsOnlyWhenRunning
    group_1 : T_SafeGroup;
    fb_1 : T_SafeDecouple(group := group_1);
END_VAR

Test_InputsLoopedToOutputsOnlyWhenRunning();

METHOD PRIVATE Test_InputsLoopedToOutputsOnlyWhenRunning
// note: this text did not pass the execution check against the stored diagram
StartTest(TestName := 'Test_InputsLoopedToOutputsOnlyWhenRunning');
group_1(Run := TRUE, ErrAck := FALSE); // T_SafeGroup
fb_1(DecIn3 := TRUE); // T_SafeDecouple
AssertEquals_BOOL(Expected := TRUE, Actual := fb_1.DecOut3, Message := 'input looped to output');
group_1(Run := FALSE, ErrAck := FALSE); // T_SafeGroup
fb_1(DecIn3 := TRUE); // T_SafeDecouple
AssertEquals_BOOL(Expected := FALSE, Actual := fb_1.DecOut3, Message := 'output off while the group is stopped');
FinishTest(TestName := 'Test_InputsLoopedToOutputsOnlyWhenRunning');
END_METHOD

END_FUNCTION_BLOCK

// ---- Tests/T_SafeOpMode_Tests_CFC.TcPOU
    // CFC twin of T_SafeOpMode_Tests: the same tests drawn as CFC diagrams, the way a TwinSAFE project is authored.
    FUNCTION_BLOCK T_SafeOpMode_Tests_CFC EXTENDS T_SafeCfcTestSuite
    VAR
    // Test_ExactlyOneInputSelectsOutput
    group_1 : T_SafeGroup;
    fb_1 : T_SafeOpMode(group := group_1);
    // Test_ConnectedRestartRequiresRestartSequence
    group_2 : T_SafeGroup;
    fb_2 : T_SafeOpMode(group := group_2);
    // Test_SlowModeChangeGivesDiscrepancyError
    group_3 : T_SafeGroup;
    fb_3 : T_SafeOpMode(group := group_3) := (Parameters := (DiscrepancyTime := T#100MS));
    t0_3 : TON;
    t1_3 : TON;
    trig1_3 : R_TRIG;
END_VAR

Test_ExactlyOneInputSelectsOutput();
Test_ConnectedRestartRequiresRestartSequence();
Test_SlowModeChangeGivesDiscrepancyError();

METHOD PRIVATE Test_ExactlyOneInputSelectsOutput
// note: this text did not pass the execution check against the stored diagram
StartTest(TestName := 'Test_ExactlyOneInputSelectsOutput');
group_1(Run := TRUE, ErrAck := FALSE); // T_SafeGroup
fb_1(OpIn1 := FALSE, OpIn2 := TRUE); // T_SafeOpMode
group_1(Run := TRUE, ErrAck := FALSE); // T_SafeGroup
fb_1(OpIn1 := FALSE, OpIn2 := TRUE); // T_SafeOpMode
AssertEquals_BOOL(Expected := TRUE, Actual := fb_1.OpOut2, Message := 'selected mode output on');
AssertEquals_BOOL(Expected := FALSE, Actual := fb_1.OpOut1, Message := 'other outputs off');
AssertEquals_BYTE(Expected := TO_BYTE(E_SafeFbState.Run), Actual := fb_1.State, Message := 'state RUN');
group_1(Run := TRUE, ErrAck := FALSE); // T_SafeGroup
fb_1(OpIn1 := TRUE, OpIn2 := TRUE); // T_SafeOpMode
AssertEquals_BOOL(Expected := FALSE, Actual := fb_1.OpOut2, Message := 'all outputs off with two modes selected');
AssertEquals_BYTE(Expected := TO_BYTE(E_SafeFbState.Safe), Actual := fb_1.State, Message := 'state SAFE');
FinishTest(TestName := 'Test_ExactlyOneInputSelectsOutput');
END_METHOD

METHOD PRIVATE Test_ConnectedRestartRequiresRestartSequence
// note: this text did not pass the execution check against the stored diagram
StartTest(TestName := 'Test_ConnectedRestartRequiresRestartSequence');
group_2(Run := TRUE, ErrAck := FALSE); // T_SafeGroup
fb_2(Restart := FALSE, OpIn1 := TRUE, OpIn2 := FALSE); // T_SafeOpMode
group_2(Run := TRUE, ErrAck := FALSE); // T_SafeGroup
fb_2(Restart := FALSE, OpIn1 := TRUE, OpIn2 := FALSE); // T_SafeOpMode
AssertEquals_BOOL(Expected := FALSE, Actual := fb_2.OpOut1, Message := 'no output before restart');
group_2(Run := TRUE, ErrAck := FALSE); // T_SafeGroup
fb_2(Restart := TRUE, OpIn1 := TRUE, OpIn2 := FALSE); // T_SafeOpMode
AssertEquals_BYTE(Expected := TO_BYTE(E_SafeFbState.Start), Actual := fb_2.State, Message := 'state START while restart held');
group_2(Run := TRUE, ErrAck := FALSE); // T_SafeGroup
fb_2(Restart := FALSE, OpIn1 := TRUE, OpIn2 := FALSE); // T_SafeOpMode
AssertEquals_BOOL(Expected := TRUE, Actual := fb_2.OpOut1, Message := 'output on after restart falling edge');
FinishTest(TestName := 'Test_ConnectedRestartRequiresRestartSequence');
END_METHOD

METHOD PRIVATE Test_SlowModeChangeGivesDiscrepancyError
// note: this text did not pass the execution check against the stored diagram
StartTest(TestName := 'Test_SlowModeChangeGivesDiscrepancyError');
t0_3(IN := TRUE, PT := T#20MS); // TON
t1_3(IN := TRUE, PT := T#250MS); // TON
trig1_3(CLK := t1_3.Q); // R_TRIG
group_3(Run := TRUE, ErrAck := FALSE); // T_SafeGroup
fb_3(OpIn1 := NOT t0_3.Q, OpIn2 := FALSE); // T_SafeOpMode
IF trig1_3.Q THEN AssertEquals_BOOL(Expected := TRUE, Actual := fb_3.Error, Message := 'discrepancy error after time without a mode'); END_IF
IF trig1_3.Q THEN AssertEquals_BYTE(Expected := TO_BYTE(E_SafeFbState.Error), Actual := fb_3.State, Message := 'state ERROR'); END_IF
IF trig1_3.Q THEN AssertEquals_WORD(Expected := WORD#1, Actual := fb_3.Diag, Message := 'diag bit 0'); END_IF
IF trig1_3.Q THEN FinishTest(TestName := 'Test_SlowModeChangeGivesDiscrepancyError'); END_IF
END_METHOD

END_FUNCTION_BLOCK

// ---- Tests/T_SafeRs_Tests_CFC.TcPOU
    // CFC twin of T_SafeRs_Tests: the same tests drawn as CFC diagrams, the way a TwinSAFE project is authored.
    FUNCTION_BLOCK T_SafeRs_Tests_CFC EXTENDS T_SafeCfcTestSuite
    VAR
    // Test_ResetDominantLatch
    group_1 : T_SafeGroup;
    fb_1 : T_SafeRs(group := group_1);
END_VAR

Test_ResetDominantLatch();

METHOD PRIVATE Test_ResetDominantLatch
// note: this text did not pass the execution check against the stored diagram
StartTest(TestName := 'Test_ResetDominantLatch');
group_1(Run := TRUE, ErrAck := FALSE); // T_SafeGroup
fb_1(Set := TRUE, Reset := FALSE); // T_SafeRs
AssertEquals_BOOL(Expected := TRUE, Actual := fb_1.RsOut, Message := 'set');
fb_1(Set := FALSE, Reset := FALSE); // T_SafeRs
AssertEquals_BOOL(Expected := TRUE, Actual := fb_1.RsOut, Message := 'held');
fb_1(Set := TRUE, Reset := TRUE); // T_SafeRs
AssertEquals_BOOL(Expected := FALSE, Actual := fb_1.RsOut, Message := 'reset dominant');
FinishTest(TestName := 'Test_ResetDominantLatch');
END_METHOD

END_FUNCTION_BLOCK

// ---- Tests/T_SafeSr_Tests_CFC.TcPOU
    // CFC twin of T_SafeSr_Tests: the same tests drawn as CFC diagrams, the way a TwinSAFE project is authored.
    FUNCTION_BLOCK T_SafeSr_Tests_CFC EXTENDS T_SafeCfcTestSuite
    VAR
    // Test_SetDominantLatch
    group_1 : T_SafeGroup;
    fb_1 : T_SafeSr(group := group_1);
END_VAR

Test_SetDominantLatch();

METHOD PRIVATE Test_SetDominantLatch
// note: this text did not pass the execution check against the stored diagram
StartTest(TestName := 'Test_SetDominantLatch');
group_1(Run := TRUE, ErrAck := FALSE); // T_SafeGroup
fb_1(Set := TRUE, Reset := TRUE); // T_SafeSr
AssertEquals_BOOL(Expected := TRUE, Actual := fb_1.SrOut, Message := 'set dominant');
fb_1(Set := FALSE, Reset := TRUE); // T_SafeSr
AssertEquals_BOOL(Expected := FALSE, Actual := fb_1.SrOut, Message := 'reset');
fb_1(Set := FALSE, Reset := FALSE); // T_SafeSr
AssertEquals_BOOL(Expected := FALSE, Actual := fb_1.SrOut, Message := 'held');
FinishTest(TestName := 'Test_SetDominantLatch');
END_METHOD

END_FUNCTION_BLOCK

// ---- Tests/T_SafeTon_Tests_CFC.TcPOU
    // CFC twin of T_SafeTon_Tests: the same tests drawn as CFC diagrams, the way a TwinSAFE project is authored.
    FUNCTION_BLOCK T_SafeTon_Tests_CFC EXTENDS T_SafeCfcTestSuite
    VAR
    // Test_OutputDelayedOn
    group_1 : T_SafeGroup;
    fb_1 : T_SafeTon(group := group_1) := (Parameters := (DelayTime := T#100MS));
    trigStart_1 : R_TRIG;
    t1_1 : TON;
    trig1_1 : R_TRIG;
END_VAR

Test_OutputDelayedOn();

METHOD PRIVATE Test_OutputDelayedOn
// note: this text did not pass the execution check against the stored diagram
